(* IEC 61131-3 sources: plc-iiot-stack/src/Interfaces/I_MqttClient, 4 files *)

(* ---- Connect.method.decl.st ---- *)
// Запросить подключение к брокеру с параметрами stCfg (включая LWT). TRUE — запрос принят;
// подключение состоялось, когда IsConnected() = TRUE.
METHOD Connect : BOOL
VAR_IN_OUT CONSTANT
    // lint:allow STL007 параметр VAR_IN_OUT CONSTANT — ссылка только для чтения, а не константа
    stCfg : ST_MqttBrokerCfg;
END_VAR

(* ---- Publish.method.decl.st ---- *)
// Поставить сообщение в очередь публикации. TRUE — клиент принял сообщение (есть связь и место в очереди);
// FALSE — не принял, вызывающий повторит позже.
METHOD Publish : BOOL
VAR_INPUT
    sTopic : STRING(GVL_Const.MQTT_TOPIC_LEN);
    eQos : E_MqttQos;
    xRetain : BOOL;
END_VAR
VAR_IN_OUT CONSTANT
    // lint:allow STL007 параметр VAR_IN_OUT CONSTANT — ссылка только для чтения, а не константа
    sPayload : STRING(GVL_Const.MQTT_PAYLOAD_LEN);
END_VAR

(* ---- Receive.method.decl.st ---- *)
// Забрать одно принятое сообщение из очереди клиента. TRUE — сообщение есть (sTopic и sPayload заполнены);
// xTruncated — текст длиннее буфера sPayload и обрезан; xRetained — сообщение пришло с флагом retain.
METHOD Receive : BOOL
VAR_IN_OUT
    sTopic : STRING(GVL_Const.MQTT_TOPIC_LEN);
    sPayload : STRING(GVL_Const.MQTT_CMD_PAYLOAD_LEN);
END_VAR
VAR_OUTPUT
    xTruncated : BOOL;
    xRetained : BOOL;
END_VAR

(* ---- Subscribe.method.decl.st ---- *)
// Подписаться на фильтр топиков (допустимы + и #). TRUE — запрос подписки принят.
METHOD Subscribe : BOOL
VAR_INPUT
    sTopicFilter : STRING(GVL_Const.MQTT_TOPIC_LEN);
    eQos : E_MqttQos;
END_VAR
